# EPICS autosave request: iocs/ad/csimdetector-ioc/db/ADCSimDetectorN_settings.req
$(P)$(R)Amplitude
$(P)$(R)Offset
$(P)$(R)Period
$(P)$(R)Phase
$(P)$(R)Noise
